RoboDK station: UR5_CB3.rdk

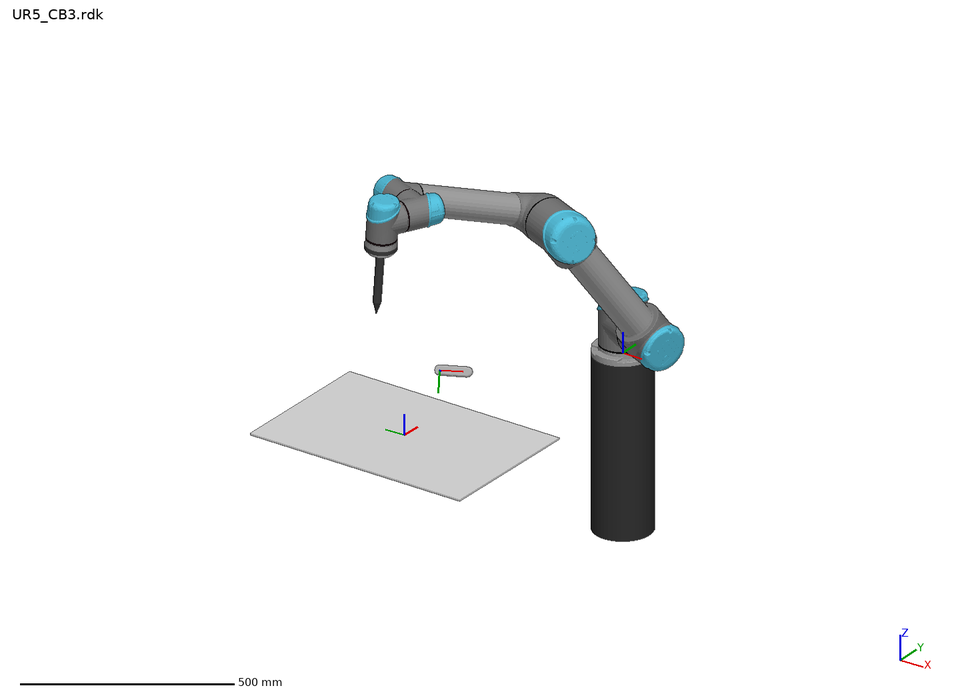
[picture v0: the station drawn from its stored meshes, robots at their saved joint values, targets as dots, program paths as lines]
Station diplomski (saved by RoboDK 5.9.0). Poses are relative to the parent item; angles as X-Y-Z fixed-axis rotations.
  - frame UR5 Base at (0, 0, 0) mm
    - robot UR5: 6 axes
        modified DH rows (alpha deg, a mm, theta deg, d mm): 0, 0, 0, 89.2; 90, 0, 180, 0; 0, 425, 0, 0; 0, 392, 0, 109.3; -90, 0, 0, 94.75; 90, 0, 180, 82.5
        joint limits [-360, -360, -360, -360, -360, -360] to [360, 360, 360, 360, 360, 360]; home [0, -90, -90, 0, 90, 0]; saved at [65.4, -54.37, 35.32, -71.74, -95.46, 1.64]
      - tool Zivid Pointed Hand-Eye Verification Tool, TCP at (0, 0, 290) mm, size 79 x 79 x 190 mm
  - frame ploca_frame at (-166.19, -648.49, -1.03) mm, rotated rx 0.22 ry -0.24 rz 89.53 deg
    - object ploca at (0, 0, 0) mm, rotated rx 0 ry 0 rz 90 deg, size 600 x 400 x 4.4 mm, geometry from Cube-100mm.sld
  - frame camera_frame at (460.57, -1399.89, 643.51) mm, rotated rx -118.2 ry 2.2 rz 30.15 deg
    - object Intel RealSense D435 Camera at (0, 0, 0) mm, size 89.8 x 25 x 25.1 mm, geometry from Intel-RealSense-D435-Camera.sld
  - object Cylinder 50x150mm at (0, 0, -452) mm, size 150 x 150 x 450 mm, geometry from Cylinder-50x150mm.sld
  - Python program Provjera (listed below)
  - Python program Robot_kamera_snap (listed below)
  - Python program Kamera_ploca_real (listed below)

--- Python program Provjera ---
from robodk import robolink, robomath
import math
import time

def provjeri_kontinuirano_crtanje_animirano(animate=True):
    RDK = robolink.Robolink()

    # 1. Dohvaćanje robota i alata
    robot = RDK.ItemUserPick(
        'Odaberi UR5 robota',
        robolink.ITEM_TYPE_ROBOT
    )

    if not robot.Valid():
        print("Robot nije odabran.")
        return

    tool = robot.Childs()[0] if robot.Childs() else None
    if not tool:
        print("UPOZORENJE: Robot nema pričvršćen alat!")
        return

    robot.setTool(tool)
    print(f"Aktivan alat: {tool.Name()}")

    # Odabir frame-a ploče
    board_frame = RDK.ItemUserPick(
        'Odaberi Frame od Bijele Ploče',
        robolink.ITEM_TYPE_FRAME
    )

    if not board_frame.Valid():
        print("Frame ploče nije odabran.")
        return

    # 2. Dimenzije ploče i parametri crtanja
    SIRINA = 550            # mm, lokalna Y os ploče
    VISINA = 350            # mm, lokalna X os ploče
    KORAK = 10              # mm, razmak točaka za IK provjeru
    RAZMAK_LINIJA = 50      # mm, vertikalni razmak horizontalnih linija

    # Orijentacija alata: TCP gleda prema ploči
    orijentacija_alata = robomath.rotx(math.pi)

    # ------------------------------------------------------------------
    # IZRAČUN DINAMIČKOG KUTA PRVOG ZGLOBA (J1) PREMA -X OSI PLOČE
    # ------------------------------------------------------------------
    # Dohvaćanje poze ploče u odnosu na bazu robota
    pose_board_rel = robot.PoseAbs().inv() * board_frame.PoseAbs()

    # Ekstrakcija X-osi ploče (vektora) u koordinatnom sustavu robota
    vx = pose_board_rel.VX()

    # Prema novoj logici promatramo -X os ploče
    neg_vx = [-vx[0], -vx[1], -vx[2]]

    # Izračun kuta između X-osi baze robota (1,0,0) i -X osi ploče u XY ravnini.
    # atan2 vraća + za CCW (suprotno od kazaljke) i - za CW (u smjeru kazaljke)
    kut_relativni_rad = math.atan2(neg_vx[1], neg_vx[0])
    kut_relativni_deg = math.degrees(kut_relativni_rad)

    # J1 je baznih -50 + relativni kut
    j1_target = -50 + kut_relativni_deg

    # Normalizacija kuta na raspon [-180, 180] radi urednije rotacije zgloba
    while j1_target > 180:
        j1_target -= 360
    while j1_target <= -180:
        j1_target += 360

    print(f"Kut -X osi ploče u odnosu na X os baze: {kut_relativni_deg:.2f}°")
    print(f"Dinamički postavljen J1: {j1_target:.2f}°")

    # Postavljanje robota u zadanu POČETNU KONFIGURACIJU s izračunatim J1
    J_POCETNI = [j1_target, -90, -105, -60, 90, 0]

    print(f"Putujem u početnu (Home) poziciju MoveJ kretnjom: {J_POCETNI}...")

    # Korištenje isključivo MoveJ kretnje za odlazak u Home poziciju
    try:
        robot.setPoseFrame(robot.Parent()) # Osiguraj da smo u bazi robota
        robot.MoveJ(J_POCETNI)
        print("Robot je uspješno stigao u početnu konfiguraciju.")
    except Exception as e:
        print(f"Greška pri odlasku u Home poziciju: {e}")
        return

    tcp_pose = robot.PoseTool()

    uspjesne_horizontalne = 0
    uspjesni_vertikalni_pomaci = 0
    putanja_moguca = True

    # Kada nije animirano, RoboDK ne osvježava 3D prikaz.
    if not animate:
        RDK.Render(False)

    print(f"Započinjem provjeru kontinuirane putanje po ploči "
          f"{SIRINA} x {VISINA} mm...")
    print(f"Animacija: {'UKLJUČENA' if animate else 'ISKLJUČENA'}")

    try:
        # Kretanje po X osi ploče: od donjeg prema gornjem dijelu
        x_vrijednosti = list(
            range(
                int(-VISINA / 2),
                int(VISINA / 2) + 1,
                RAZMAK_LINIJA
            )
        )

        if x_vrijednosti[-1] != int(VISINA / 2):
            x_vrijednosti.append(int(VISINA / 2))

        # Robot prvo ide s desne na lijevu stranu.
        smjer_desno_prema_lijevo = True

        zadnji_j_list = list(J_POCETNI)
        prva_tocka_putanje = True

        for indeks_linije, x_visina in enumerate(x_vrijednosti):

            if smjer_desno_prema_lijevo:
                y_vrijednosti = list(
                    range(
                        int(SIRINA / 2),
                        int(-SIRINA / 2) - 1,
                        -KORAK
                    )
                )
                smjer_teksta = "desno -> lijevo"
            else:
                y_vrijednosti = list(
                    range(
                        int(-SIRINA / 2),
                        int(SIRINA / 2) + 1,
                        KORAK
                    )
                )
                smjer_teksta = "lijevo -> desno"

            zavrsni_y = int(-SIRINA / 2) if smjer_desno_prema_lijevo else int(SIRINA / 2)
            if y_vrijednosti[-1] != zavrsni_y:
                y_vrijednosti.append(zavrsni_y)

            print(f"Provjera horizontalne linije X={x_visina} mm ({smjer_teksta})")

            # ----------------------------------------------------------
            # HORIZONTALNI DIO PUTANJE
            # ----------------------------------------------------------
            for y_sirina in y_vrijednosti:

                poza_lokalno = (
                    robomath.transl(x_visina, y_sirina, 0)
                    * orijentacija_alata
                )

                poza_apsolutno = board_frame.PoseAbs() * poza_lokalno
                poza_u_bazi_robota = (
                    robot.PoseAbs().inv() * poza_apsolutno
                )

                # Prilaz PRVOJ točci pomoću MoveJ i MoveL
                if prva_tocka_putanje:
                    print("-" * 40)
                    print("Prilazak prvoj točci (Z=100mm offset uz MoveJ, pa MoveL na ploču)...")

                    # Kreiranje offset poze 100mm iznad ploče (po Z osi ploče)
                    poza_lokalno_offset = (
                        robomath.transl(x_visina, y_sirina, 100)
                        * orijentacija_alata
                    )
                    poza_apsolutno_offset = board_frame.PoseAbs() * poza_lokalno_offset
                    poza_u_bazi_robota_offset = robot.PoseAbs().inv() * poza_apsolutno_offset

                    try:
                        # Osiguraj da se kretnje računaju u odnosu na bazu robota
                        robot.setPoseFrame(robot.Parent())

                        # Brzi pomak iznad prve točke
                        robot.MoveJ(poza_u_bazi_robota_offset)
                        # Linearno spuštanje vrha alata na ploču
                        robot.MoveL(poza_u_bazi_robota)

                        # Ažuriraj zglobove nakon pomaka kako bi se nastavila ručna IK provjera koda
                        zadnji_j = robot.Joints().list()
                        zadnji_j_list = zadnji_j
                        prva_tocka_putanje = False

                        print("Prilaz uspješan! Započinjem crtanje.")
                        print("-" * 40)
                        continue # Prelazi na prvu točku crtanja
                    except Exception as e:
                        print(f"PUTANJA PALA: Greška pri inicijalnom prilazu: {e}")
                        putanja_moguca = False
                        break

                # Redovno crtanje s manualnom provjerom IK i glatkoće za animaciju
                trenutni_zglobovi = robot.SolveIK(
                    poza_u_bazi_robota,
                    zadnji_j_list,
                    tcp_pose
                )
                trenutni_j_list = trenutni_zglobovi.list()

                if len(trenutni_j_list) != 6:
                    print(
                        f"PUTANJA PALA: IK ne postoji na "
                        f"X={x_visina}, Y={y_sirina} mm."
                    )
                    putanja_moguca = False
                    break

                for i in range(6):
                    razlika_kuta = abs(
                        trenutni_j_list[i] - zadnji_j_list[i]
                    )

                    if razlika_kuta > 15.0:
                        print(
                            f"PUTANJA PALA: trzaj na "
                            f"X={x_visina}, Y={y_sirina} mm "
                            f"(zglob {i + 1}: {razlika_kuta:.2f}°)."
                        )
                        putanja_moguca = False
                        break

                if not putanja_moguca:
                    break

                robot.setJoints(trenutni_j_list)
                if animate:
                    time.sleep(0.02)

                if RDK.Collisions() > 0:
                    print(
                        f"PUTANJA PALA: sudar na "
                        f"X={x_visina}, Y={y_sirina} mm."
                    )
                    putanja_moguca = False
                    break

                zadnji_j_list = trenutni_j_list

            if not putanja_moguca:
                break

            uspjesne_horizontalne += 1

            # ----------------------------------------------------------
            # VERTIKALNI DIO PUTANJE
            # ----------------------------------------------------------
            if indeks_linije < len(x_vrijednosti) - 1:
                sljedeci_x = x_vrijednosti[indeks_linije + 1]
                rubni_y = zavrsni_y
                korak_x = KORAK if sljedeci_x > x_visina else -KORAK

                x_vertikalne_tocke = list(
                    range(
                        x_visina + korak_x,
                        sljedeci_x + korak_x,
                        korak_x
                    )
                )

                x_vertikalne_tocke = [
                    x for x in x_vertikalne_tocke
                    if (
                        x <= sljedeci_x
                        if korak_x > 0
                        else x >= sljedeci_x
                    )
                ]

                if not x_vertikalne_tocke or x_vertikalne_tocke[-1] != sljedeci_x:
                    x_vertikalne_tocke.append(sljedeci_x)

                print(
                    f"Provjera vertikalnog prijelaza: "
                    f"X={x_visina} -> X={sljedeci_x} mm, "
                    f"Y={rubni_y} mm"
                )

                for x_vertikalno in x_vertikalne_tocke:

                    poza_lokalno = (
                        robomath.transl(x_vertikalno, rubni_y, 0)
                        * orijentacija_alata
                    )

                    poza_apsolutno = board_frame.PoseAbs() * poza_lokalno
                    poza_u_bazi_robota = (
                        robot.PoseAbs().inv() * poza_apsolutno
                    )

                    trenutni_zglobovi = robot.SolveIK(
                        poza_u_bazi_robota,
                        zadnji_j_list,
                        tcp_pose
                    )
                    trenutni_j_list = trenutni_zglobovi.list()

                    if len(trenutni_j_list) != 6:
                        print(
                            f"PUTANJA PALA: IK ne postoji na "
                            f"vertikalnom dijelu "
                            f"X={x_vertikalno}, Y={rubni_y} mm."
                        )
                        putanja_moguca = False
                        break

                    for i in range(6):
                        razlika_kuta = abs(
                            trenutni_j_list[i] - zadnji_j_list[i]
                        )

                        if razlika_kuta > 15.0:
                            print(
                                f"PUTANJA PALA: trzaj na vertikalnom dijelu "
                                f"X={x_vertikalno}, Y={rubni_y} mm "
                                f"(zglob {i + 1}: {razlika_kuta:.2f}°)."
                            )
                            putanja_moguca = False
                            break

                    if not putanja_moguca:
                        break

                    robot.setJoints(trenutni_j_list)

                    if animate:
                        time.sleep(0.02)

                    if RDK.Collisions() > 0:
                        print(
                            f"PUTANJA PALA: sudar na vertikalnom dijelu "
                            f"X={x_vertikalno}, Y={rubni_y} mm."
                        )
                        putanja_moguca = False
                        break

                    zadnji_j_list = trenutni_j_list

                if not putanja_moguca:
                    break

                uspjesni_vertikalni_pomaci += 1

            smjer_desno_prema_lijevo = not smjer_desno_prema_lijevo

    finally:
        if not animate:
            RDK.Render(True)

    print("-" * 55)
    print("REZULTAT PROVJERE KONTINUIRANOG CRTANJA:")

    if putanja_moguca:
        print("STATUS: CIJELA KONTINUIRANA PUTANJA JE MOGUĆA.")
    else:
        print("STATUS: PUTANJA JE PREKINUTA ZBOG IK-a, TRZAJA ILI SUDARA.")

    print(f"Uspješno nacrtanih horizontalnih linija: {uspjesne_horizontalne}")
    print(f"Uspješno provjerenih vertikalnih prijelaza: {uspjesni_vertikalni_pomaci}")
    print("-" * 55)

if __name__ == '__main__':
    provjeri_kontinuirano_crtanje_animirano(animate=True)

--- Python program Robot_kamera_snap ---
from robodk import robolink, robomath
import numpy as np
import os
import socket
import struct
import math

def get_current_joints(robot_ip):
    """
    Spaja se na UR Real-Time port (30003), čita paket i izvlači
    stvarne pozicije zglobova (q_actual) te ih vraća u stupnjevima.
    """
    port = 30003
    try:
        s = socket.socket(socket.AF_INET, socket.SOCK_STREAM)
        s.settimeout(2.0)
        s.connect((robot_ip, port))

        # Čitamo barem 300 byteova jer se q_actual nalazi na offsetu 252
        packet = b''
        while len(packet) < 300:
            chunk = s.recv(4096)
            if not chunk:
                break
            packet += chunk
        s.close()

        if len(packet) >= 300:
            # U UR paketu (CB3 i e-Series), 'q_actual' kreće od 252. bytea.
            # Format je 6 double vrijednosti (8 byteova svaka), Big-Endian (!6d)
            joints_rad = struct.unpack('!6d', packet[252:300])

            # RoboDK koristi stupnjeve, pa radijane pretvaramo u stupnjeve
            joints_deg = [math.degrees(j) for j in joints_rad]
            return joints_deg
        else:
            print("GREŠKA: Nije primljeno dovoljno podataka s robota.")
            return None

    except Exception as e:
        print(f"GREŠKA pri spajanju na fizičkog robota: {e}")
        return None

def main():
    # 1. Spajanje na aktivnu RoboDK instancu
    RDK = robolink.Robolink()

    # 2. Pronalazak frame-ova u postaji
    frame_board = RDK.Item('UR5e Base', robolink.ITEM_TYPE_FRAME)
    frame_camera = RDK.Item('camera_frame', robolink.ITEM_TYPE_FRAME)

    # Pronalazak robota (Provjeri je li ime točno onako kako piše u stablu postaje!)
    robot = RDK.Item('UR5e', robolink.ITEM_TYPE_ROBOT)

    # Provjera jesu li objekti ispravno pronađeni
    if not frame_board.Valid():
        print("GREŠKA: Frame 'UR5e Base' nije pronađen u postaji!")
        return
    if not frame_camera.Valid():
        print("GREŠKA: Frame 'camera_frame' nije pronađen u postaji!")
        return
    if not robot.Valid():
        print("GREŠKA: Robot 'UR5e' nije pronađen u postaji! Provjeri točno ime u stablu.")
        return

    # 3. Učitavanje matrice iz .npy datoteke
    path_to_matrix = r"C:/Users/User/PycharmProjects/Diplomski_realsense/kalibracija_res/T_base_cam.npy"

    if not os.path.exists(path_to_matrix):
        print(f"GREŠKA: Datoteka {path_to_matrix} ne postoji.")
        return

    T_cam_board_np = np.load(path_to_matrix)

    # 4. Pretvorba OpenCV numpy 4x4 matrice u RoboDK Mat objekt
    pose_cam_rel_board = robomath.Mat(T_cam_board_np.tolist())

    # 5. Izračun i primjena nove pozicije
    pose_board_abs = frame_board.PoseAbs()
    pose_camera_abs = pose_board_abs * pose_cam_rel_board
    frame_camera.setPoseAbs(pose_camera_abs)
    print("Uspješno! 'camera_frame' je pomaknut na točnu poziciju.")

    # 6. Dohvaćanje pozicije zglobova s fizičkog robota i snap u RoboDK
    robot_ip = "192.168.40.18"
    print(f"Dohvaćam poziciju zglobova s IP adrese {robot_ip}...")

    joints_deg = get_current_joints(robot_ip)
    if joints_deg:
        # Postavljamo virtualnog robota u izračunate kuteve
        robot.setJoints(joints_deg)
        print(f"Virtualni robot sinkroniziran s fizičkim. Kutevi: {[round(j, 2) for j in joints_deg]}")
    else:
        print("Prekid sinkronizacije: nije uspjelo čitanje s fizičkog robota.")

if __name__ == "__main__":
    main()

--- Python program Kamera_ploca_real ---
from robodk import robolink, robomath
import numpy as np
import os

def main():
    # 1. Spajanje na aktivnu RoboDK instancu
    RDK = robolink.Robolink()

    # 2. Pronalazak frame-ova u postaji
    frame_board = RDK.Item('ploca_frame', robolink.ITEM_TYPE_FRAME)
    frame_camera = RDK.Item('camera_frame', robolink.ITEM_TYPE_FRAME)

    # Provjera jesu li frame-ovi ispravno pronađeni
    if not frame_board.Valid():
        print("GREŠKA: Frame 'ploca_frame' nije pronađen u postaji!")
        return
    if not frame_camera.Valid():
        print("GREŠKA: Frame 'camera_frame' nije pronađen u postaji!")
        return

    # 3. Učitavanje matrice iz .npy datoteke
    # Koristimo matricu T_cam_board koja opisuje poziciju ploče u odnosu na kameru
    path_to_matrix = r"C:/Users/User/PycharmProjects/Diplomski_realsense/kalibracija_res/T_cam_board.npy"

    if not os.path.exists(path_to_matrix):
        print(f"GREŠKA: Datoteka {path_to_matrix} ne postoji.")
        return

    T_board_rel_cam_np = np.load(path_to_matrix)

    # 4. Pretvorba OpenCV numpy 4x4 matrice u RoboDK Mat objekt
    pose_board_rel_cam = robomath.Mat(T_board_rel_cam_np.tolist())

    # 5. Izračun i primjena nove pozicije
    # Dohvaćamo apsolutnu poziciju kamere u postaji (koja sada ostaje fiksna)
    pose_camera_abs = frame_camera.PoseAbs()

    # Apsolutna pozicija ploče = Aps. pozicija kamere * Relativna pozicija ploče (u odnosu na kameru)
    pose_board_abs = pose_camera_abs * pose_board_rel_cam

    # Postavljamo novu apsolutnu poziciju ploče, a camera_frame ostaje netaknut!
    frame_board.setPoseAbs(pose_board_abs)

    print("Uspješno! 'ploca_frame' je pomaknut na točnu poziciju u odnosu na fiksni 'camera_frame'.")

if __name__ == "__main__":
    main()
